Fanuc KAREL source: KT00742.KL

PROGRAM KT00742
%NOLOCKGROUP
VAR
  ARG: ARRAY[4] OF VECTOR
  OUT: BOOLEAN
BEGIN
  OUT = UNINIT(ARG)
END KT00742
